Staubli VAL3: pointMove.pgx

public program pointMove(string x_sKey, num x_nIndex)
  local num l_nType
  local frame l_fFrame
  local pointRx l_pPoint
  local tool l_tTool
  local jointRx l_jJoint
  local bool l_bResult
  local jointRx l_jHere
  local pointRx l_pPoint1
  local num l_nSigIndex
  local bool l_bSigValue
  local num l_nSigValue
  local bool l_bErr
begin
  link(l_fFrame,world)
  link(l_tTool,flange)
  //link(l_pPoint,world)
  l_nType=trajTemp:tTrajItem[x_sKey].pPointItem[x_nIndex].pParaItem.nMoveType
  call savedata:getFrame(trajTemp:tTrajItem[x_sKey].nFrameIndex,l_fFrame)
  call savedata:getTool(trajTemp:tTrajItem[x_sKey].nToolIndex,l_tTool)
  link(l_pPoint,l_fFrame)
  link(l_pPoint1,l_fFrame)
  l_pPoint.trsf=trajTemp:tTrajItem[x_sKey].pPointItem[x_nIndex].pPointRx.trsf
  l_pPoint.config=trajTemp:tTrajItem[x_sKey].pPointItem[x_nIndex].pPointRx.config
  l_pPoint1.trsf=trajTemp:tTrajItem[x_sKey].pPointItem[x_nIndex].pInter.trsf
  l_pPoint1.config=trajTemp:tTrajItem[x_sKey].pPointItem[x_nIndex].pInter.config
  l_jJoint=trajTemp:tTrajItem[x_sKey].pPointItem[x_nIndex].jJointRx
  l_nSigIndex=trajTemp:tTrajItem[x_sKey].pPointItem[x_nIndex].pParaItem.nActionIndex
  l_bSigValue=(trajTemp:tTrajItem[x_sKey].pPointItem[x_nIndex].pParaItem.nSigValue!=0)
  l_nSigValue=trajTemp:tTrajItem[x_sKey].pPointItem[x_nIndex].pParaItem.nSigValue
  if rs:_nOmacStat==9 and workingMode()==1 and isPowered()
    // if !isEmpty()
    stopMove()
    resetMotion()
    l_jHere=herej()
    movej(l_jHere,flange,mSim)
    // endIf
    switch l_nType
      case 1
        call isPointOK(x_sKey,x_nIndex,l_bResult)
        if l_bResult
          movel(l_pPoint,l_tTool,mSim)
        endIf
      break
      case 0
        movej(l_jJoint,l_tTool,mSim)
      break
      case 2
        movec(l_pPoint1,l_pPoint,l_tTool,mSim)
      break
      //Add by Liu Zhengang 20251028
      case 3
        //dIn
        waitEndMove()
        if watch($isKeyPressed(14),5)==true
          call io:waitDigInput(io:dInput[l_nSigIndex],l_bSigValue,l_bErr)
          popUpMsg("din"+"["+toString("",l_nSigIndex)+"]"+"执行成功")
        endIf

      break
      case 4
        //dOut
        waitEndMove()
        if watch($isKeyPressed(14),5)==true

          call io:setDigOutput(io:dOutput[l_nSigIndex],l_bSigValue,l_bErr)
          popUpMsg("dout"+"["+toString("",l_nSigIndex)+"]"+"执行成功")
        endIf
      break
      case 5
        //ain
        waitEndMove()
        if watch($isKeyPressed(14),5)==true
          call io:waitAnaInput(io:aInput[l_nSigIndex],l_nSigValue,l_bErr)
          popUpMsg("ain"+"["+toString("",l_nSigIndex)+"]"+"执行成功")
        endIf

        // wait(l_nSigValue==l_nValue)
      break
      case 6
        //aout
        waitEndMove()
        if watch($isKeyPressed(14),5)==true
          call io:setAnaOutput(io:aOutput[l_nSigIndex],l_nSigValue,l_bErr)
          popUpMsg("aout"+"["+toString("",l_nSigIndex)+"]"+"执行成功")
        endIf
      break
    endSwitch
    delay(0)
  endIf
end
